(* IEC 61131-3 sources: s7-to-codesys/tests/POUs/Scenarios/FB_Totalizer_ScenarioTest, 7 files *)

(* ---- FB_Totalizer_ScenarioTest.decl.st ---- *)
// AUTO-GENERATED — не редактировать: s7conv gen-tests, сценарии scenarios/FB_Totalizer.csv
// Правка — в CSV (scenarios/README.md), затем python -m s7conv build-corpus.
// Назначение: тесты поведения сконвертированного FB_Totalizer по сценариям CSV (сценариев: 6, строк: 36):
//             один метод-тест на сценарий, строки — по порядку с моделируемым временем GVL_S7Clock.
//             Ожидаемые значения — из CSV (эталонные модели по описанию логики блока), не из
//             результата конвертации.
// Автор:      s7conv 0.1.0 (сгенерировано)
// Версия:     не указана
// Документ:   scenarios/README.md, docs/methodology.md, раздел «Проверка поведения»
FUNCTION_BLOCK FB_Totalizer_ScenarioTest EXTENDS coUnit.FB_TestSuite
VAR
    fbIntegrationAndPulses : FB_Totalizer;  // свой экземпляр на сценарий
    xIntegrationAndPulsesDone : BOOL;  // сценарий выполнен (выполняется один раз)
    fbCutoffAndEnable : FB_Totalizer;  // свой экземпляр на сценарий
    xCutoffAndEnableDone : BOOL;  // сценарий выполнен (выполняется один раз)
    fbResetLevel : FB_Totalizer;  // свой экземпляр на сценарий
    xResetLevelDone : BOOL;  // сценарий выполнен (выполняется один раз)
    fbVariableCycleTime : FB_Totalizer;  // свой экземпляр на сценарий
    xVariableCycleTimeDone : BOOL;  // сценарий выполнен (выполняется один раз)
    fbLargeStepPulsesCatchUp : FB_Totalizer;  // свой экземпляр на сценарий
    xLargeStepPulsesCatchUpDone : BOOL;  // сценарий выполнен (выполняется один раз)
    fbPulseVolumeZero : FB_Totalizer;  // свой экземпляр на сценарий
    xPulseVolumeZeroDone : BOOL;  // сценарий выполнен (выполняется один раз)
END_VAR

(* ---- CutoffAndEnable.method.impl.st ---- *)
// AUTO-GENERATED — не редактировать: scenarios/FB_Totalizer.csv, сценарий CutoffAndEnable
coUnit.TEST('CutoffAndEnable');
IF NOT xCutoffAndEnableDone THEN
    xCutoffAndEnableDone := TRUE;
    GVL_S7Clock.xSimulation := TRUE;

    // #1, t = 0 мс — 0.25 < отсечки 0.5: не считается
    GVL_S7Clock.tSimNow := T#0MS;
    fbCutoffAndEnable.flow := 0.25;
    fbCutoffAndEnable.cycleTime := T#1000MS;
    fbCutoffAndEnable.lowFlowCutoff := 0.5;
    fbCutoffAndEnable.enable := TRUE;
    fbCutoffAndEnable.reset := FALSE;
    fbCutoffAndEnable.pulseVolume := 1.0;
    fbCutoffAndEnable();
    AssertEquals_LREAL(Expected := 0.0,
                       Actual := fbCutoffAndEnable.total,
                       Delta := 0.000001,
                       Message := 'CutoffAndEnable#1 total');
    AssertEquals_LREAL(Expected := 0.0,
                       Actual := fbCutoffAndEnable.lifetimeTotal,
                       Delta := 0.000001,
                       Message := 'CutoffAndEnable#1 lifetimeTotal');
    AssertEquals_DINT(Expected := 0, Actual := fbCutoffAndEnable.pulseCount, Message := 'CutoffAndEnable#1 pulseCount');
    AssertEquals_BOOL(Expected := FALSE, Actual := fbCutoffAndEnable.pulse, Message := 'CutoffAndEnable#1 pulse');
    AssertEquals_BOOL(Expected := TRUE,
                      Actual := fbCutoffAndEnable.cutoffActive,
                      Message := 'CutoffAndEnable#1 cutoffActive');

    // #2, t = 1000 мс — обратный расход ниже отсечки: не считается
    GVL_S7Clock.tSimNow := T#1000MS;
    fbCutoffAndEnable.flow := -10.0;
    fbCutoffAndEnable();
    AssertEquals_LREAL(Expected := 0.0,
                       Actual := fbCutoffAndEnable.total,
                       Delta := 0.000001,
                       Message := 'CutoffAndEnable#2 total');
    AssertEquals_LREAL(Expected := 0.0,
                       Actual := fbCutoffAndEnable.lifetimeTotal,
                       Delta := 0.000001,
                       Message := 'CutoffAndEnable#2 lifetimeTotal');
    AssertEquals_DINT(Expected := 0, Actual := fbCutoffAndEnable.pulseCount, Message := 'CutoffAndEnable#2 pulseCount');
    AssertEquals_BOOL(Expected := FALSE, Actual := fbCutoffAndEnable.pulse, Message := 'CutoffAndEnable#2 pulse');
    AssertEquals_BOOL(Expected := TRUE,
                      Actual := fbCutoffAndEnable.cutoffActive,
                      Message := 'CutoffAndEnable#2 cutoffActive');

    // #3, t = 2000 мс — интегрирование запрещено (отсечка не активна)
    GVL_S7Clock.tSimNow := T#2000MS;
    fbCutoffAndEnable.flow := 450.0;
    fbCutoffAndEnable.enable := FALSE;
    fbCutoffAndEnable();
    AssertEquals_LREAL(Expected := 0.0,
                       Actual := fbCutoffAndEnable.total,
                       Delta := 0.000001,
                       Message := 'CutoffAndEnable#3 total');
    AssertEquals_LREAL(Expected := 0.0,
                       Actual := fbCutoffAndEnable.lifetimeTotal,
                       Delta := 0.000001,
                       Message := 'CutoffAndEnable#3 lifetimeTotal');
    AssertEquals_DINT(Expected := 0, Actual := fbCutoffAndEnable.pulseCount, Message := 'CutoffAndEnable#3 pulseCount');
    AssertEquals_BOOL(Expected := FALSE, Actual := fbCutoffAndEnable.pulse, Message := 'CutoffAndEnable#3 pulse');
    AssertEquals_BOOL(Expected := FALSE,
                      Actual := fbCutoffAndEnable.cutoffActive,
                      Message := 'CutoffAndEnable#3 cutoffActive');

    // #4, t = 3000 мс — разрешено: 0.125 м3
    GVL_S7Clock.tSimNow := T#3000MS;
    fbCutoffAndEnable.enable := TRUE;
    fbCutoffAndEnable();
    AssertEquals_LREAL(Expected := 0.125,
                       Actual := fbCutoffAndEnable.total,
                       Delta := 0.000001,
                       Message := 'CutoffAndEnable#4 total');
    AssertEquals_LREAL(Expected := 0.125,
                       Actual := fbCutoffAndEnable.lifetimeTotal,
                       Delta := 0.000001,
                       Message := 'CutoffAndEnable#4 lifetimeTotal');
    AssertEquals_DINT(Expected := 0, Actual := fbCutoffAndEnable.pulseCount, Message := 'CutoffAndEnable#4 pulseCount');
    AssertEquals_BOOL(Expected := FALSE, Actual := fbCutoffAndEnable.pulse, Message := 'CutoffAndEnable#4 pulse');
    AssertEquals_BOOL(Expected := FALSE,
                      Actual := fbCutoffAndEnable.cutoffActive,
                      Message := 'CutoffAndEnable#4 cutoffActive');

    // #5, t = 4000 мс — 0.5 = отсечке — считается: +0.5/3600 м3
    GVL_S7Clock.tSimNow := T#4000MS;
    fbCutoffAndEnable.flow := 0.5;
    fbCutoffAndEnable();
    AssertEquals_LREAL(Expected := 0.125138889,
                       Actual := fbCutoffAndEnable.total,
                       Delta := 0.000001,
                       Message := 'CutoffAndEnable#5 total');
    AssertEquals_LREAL(Expected := 0.125138889,
                       Actual := fbCutoffAndEnable.lifetimeTotal,
                       Delta := 0.000001,
                       Message := 'CutoffAndEnable#5 lifetimeTotal');
    AssertEquals_DINT(Expected := 0, Actual := fbCutoffAndEnable.pulseCount, Message := 'CutoffAndEnable#5 pulseCount');
    AssertEquals_BOOL(Expected := FALSE, Actual := fbCutoffAndEnable.pulse, Message := 'CutoffAndEnable#5 pulse');
    AssertEquals_BOOL(Expected := FALSE,
                      Actual := fbCutoffAndEnable.cutoffActive,
                      Message := 'CutoffAndEnable#5 cutoffActive');

    // #6, t = 5000 мс — 0.49 < 0.5: не считается
    GVL_S7Clock.tSimNow := T#5000MS;
    fbCutoffAndEnable.flow := 0.49;
    fbCutoffAndEnable();
    AssertEquals_LREAL(Expected := 0.125138889,
                       Actual := fbCutoffAndEnable.total,
                       Delta := 0.000001,
                       Message := 'CutoffAndEnable#6 total');
    AssertEquals_LREAL(Expected := 0.125138889,
                       Actual := fbCutoffAndEnable.lifetimeTotal,
                       Delta := 0.000001,
                       Message := 'CutoffAndEnable#6 lifetimeTotal');
    AssertEquals_DINT(Expected := 0, Actual := fbCutoffAndEnable.pulseCount, Message := 'CutoffAndEnable#6 pulseCount');
    AssertEquals_BOOL(Expected := FALSE, Actual := fbCutoffAndEnable.pulse, Message := 'CutoffAndEnable#6 pulse');
    AssertEquals_BOOL(Expected := TRUE,
                      Actual := fbCutoffAndEnable.cutoffActive,
                      Message := 'CutoffAndEnable#6 cutoffActive');

    GVL_S7Clock.xSimulation := FALSE;
END_IF
coUnit.TEST_FINISHED();

(* ---- IntegrationAndPulses.method.impl.st ---- *)
// AUTO-GENERATED — не редактировать: scenarios/FB_Totalizer.csv, сценарий IntegrationAndPulses
coUnit.TEST('IntegrationAndPulses');
IF NOT xIntegrationAndPulsesDone THEN
    xIntegrationAndPulsesDone := TRUE;
    GVL_S7Clock.xSimulation := TRUE;

    // #1, t = 0 мс — 0.125 м3
    GVL_S7Clock.tSimNow := T#0MS;
    fbIntegrationAndPulses.flow := 450.0;
    fbIntegrationAndPulses.cycleTime := T#1000MS;
    fbIntegrationAndPulses.lowFlowCutoff := 0.5;
    fbIntegrationAndPulses.enable := TRUE;
    fbIntegrationAndPulses.reset := FALSE;
    fbIntegrationAndPulses.pulseVolume := 0.5;
    fbIntegrationAndPulses();
    AssertEquals_LREAL(Expected := 0.125,
                       Actual := fbIntegrationAndPulses.total,
                       Delta := 0.000001,
                       Message := 'IntegrationAndPulses#1 total');
    AssertEquals_LREAL(Expected := 0.125,
                       Actual := fbIntegrationAndPulses.lifetimeTotal,
                       Delta := 0.000001,
                       Message := 'IntegrationAndPulses#1 lifetimeTotal');
    AssertEquals_DINT(Expected := 0,
                      Actual := fbIntegrationAndPulses.pulseCount,
                      Message := 'IntegrationAndPulses#1 pulseCount');
    AssertEquals_BOOL(Expected := FALSE,
                      Actual := fbIntegrationAndPulses.pulse,
                      Message := 'IntegrationAndPulses#1 pulse');
    AssertEquals_BOOL(Expected := FALSE,
                      Actual := fbIntegrationAndPulses.cutoffActive,
                      Message := 'IntegrationAndPulses#1 cutoffActive');

    // #2, t = 1000 мс — 0.25 м3
    GVL_S7Clock.tSimNow := T#1000MS;
    fbIntegrationAndPulses();
    AssertEquals_LREAL(Expected := 0.25,
                       Actual := fbIntegrationAndPulses.total,
                       Delta := 0.000001,
                       Message := 'IntegrationAndPulses#2 total');
    AssertEquals_LREAL(Expected := 0.25,
                       Actual := fbIntegrationAndPulses.lifetimeTotal,
                       Delta := 0.000001,
                       Message := 'IntegrationAndPulses#2 lifetimeTotal');
    AssertEquals_DINT(Expected := 0,
                      Actual := fbIntegrationAndPulses.pulseCount,
                      Message := 'IntegrationAndPulses#2 pulseCount');
    AssertEquals_BOOL(Expected := FALSE,
                      Actual := fbIntegrationAndPulses.pulse,
                      Message := 'IntegrationAndPulses#2 pulse');
    AssertEquals_BOOL(Expected := FALSE,
                      Actual := fbIntegrationAndPulses.cutoffActive,
                      Message := 'IntegrationAndPulses#2 cutoffActive');

    // #3, t = 2000 мс — 0.375 м3
    GVL_S7Clock.tSimNow := T#2000MS;
    fbIntegrationAndPulses();
    AssertEquals_LREAL(Expected := 0.375,
                       Actual := fbIntegrationAndPulses.total,
                       Delta := 0.000001,
                       Message := 'IntegrationAndPulses#3 total');
    AssertEquals_LREAL(Expected := 0.375,
                       Actual := fbIntegrationAndPulses.lifetimeTotal,
                       Delta := 0.000001,
                       Message := 'IntegrationAndPulses#3 lifetimeTotal');
    AssertEquals_DINT(Expected := 0,
                      Actual := fbIntegrationAndPulses.pulseCount,
                      Message := 'IntegrationAndPulses#3 pulseCount');
    AssertEquals_BOOL(Expected := FALSE,
                      Actual := fbIntegrationAndPulses.pulse,
                      Message := 'IntegrationAndPulses#3 pulse');
    AssertEquals_BOOL(Expected := FALSE,
                      Actual := fbIntegrationAndPulses.cutoffActive,
                      Message := 'IntegrationAndPulses#3 cutoffActive');

    // #4, t = 3000 мс — 0.5 м3: импульс №1
    GVL_S7Clock.tSimNow := T#3000MS;
    fbIntegrationAndPulses();
    AssertEquals_LREAL(Expected := 0.5,
                       Actual := fbIntegrationAndPulses.total,
                       Delta := 0.000001,
                       Message := 'IntegrationAndPulses#4 total');
    AssertEquals_LREAL(Expected := 0.5,
                       Actual := fbIntegrationAndPulses.lifetimeTotal,
                       Delta := 0.000001,
                       Message := 'IntegrationAndPulses#4 lifetimeTotal');
    AssertEquals_DINT(Expected := 1,
                      Actual := fbIntegrationAndPulses.pulseCount,
                      Message := 'IntegrationAndPulses#4 pulseCount');
    AssertEquals_BOOL(Expected := TRUE,
                      Actual := fbIntegrationAndPulses.pulse,
                      Message := 'IntegrationAndPulses#4 pulse');
    AssertEquals_BOOL(Expected := FALSE,
                      Actual := fbIntegrationAndPulses.cutoffActive,
                      Message := 'IntegrationAndPulses#4 cutoffActive');

    // #5, t = 4000 мс — 0.625 м3, импульса нет
    GVL_S7Clock.tSimNow := T#4000MS;
    fbIntegrationAndPulses();
    AssertEquals_LREAL(Expected := 0.625,
                       Actual := fbIntegrationAndPulses.total,
                       Delta := 0.000001,
                       Message := 'IntegrationAndPulses#5 total');
    AssertEquals_LREAL(Expected := 0.625,
                       Actual := fbIntegrationAndPulses.lifetimeTotal,
                       Delta := 0.000001,
                       Message := 'IntegrationAndPulses#5 lifetimeTotal');
    AssertEquals_DINT(Expected := 1,
                      Actual := fbIntegrationAndPulses.pulseCount,
                      Message := 'IntegrationAndPulses#5 pulseCount');
    AssertEquals_BOOL(Expected := FALSE,
                      Actual := fbIntegrationAndPulses.pulse,
                      Message := 'IntegrationAndPulses#5 pulse');
    AssertEquals_BOOL(Expected := FALSE,
                      Actual := fbIntegrationAndPulses.cutoffActive,
                      Message := 'IntegrationAndPulses#5 cutoffActive');

    // #6, t = 5000 мс — 0.75 м3
    GVL_S7Clock.tSimNow := T#5000MS;
    fbIntegrationAndPulses();
    AssertEquals_LREAL(Expected := 0.75,
                       Actual := fbIntegrationAndPulses.total,
                       Delta := 0.000001,
                       Message := 'IntegrationAndPulses#6 total');
    AssertEquals_LREAL(Expected := 0.75,
                       Actual := fbIntegrationAndPulses.lifetimeTotal,
                       Delta := 0.000001,
                       Message := 'IntegrationAndPulses#6 lifetimeTotal');
    AssertEquals_DINT(Expected := 1,
                      Actual := fbIntegrationAndPulses.pulseCount,
                      Message := 'IntegrationAndPulses#6 pulseCount');
    AssertEquals_BOOL(Expected := FALSE,
                      Actual := fbIntegrationAndPulses.pulse,
                      Message := 'IntegrationAndPulses#6 pulse');
    AssertEquals_BOOL(Expected := FALSE,
                      Actual := fbIntegrationAndPulses.cutoffActive,
                      Message := 'IntegrationAndPulses#6 cutoffActive');

    // #7, t = 6000 мс — 0.875 м3
    GVL_S7Clock.tSimNow := T#6000MS;
    fbIntegrationAndPulses();
    AssertEquals_LREAL(Expected := 0.875,
                       Actual := fbIntegrationAndPulses.total,
                       Delta := 0.000001,
                       Message := 'IntegrationAndPulses#7 total');
    AssertEquals_LREAL(Expected := 0.875,
                       Actual := fbIntegrationAndPulses.lifetimeTotal,
                       Delta := 0.000001,
                       Message := 'IntegrationAndPulses#7 lifetimeTotal');
    AssertEquals_DINT(Expected := 1,
                      Actual := fbIntegrationAndPulses.pulseCount,
                      Message := 'IntegrationAndPulses#7 pulseCount');
    AssertEquals_BOOL(Expected := FALSE,
                      Actual := fbIntegrationAndPulses.pulse,
                      Message := 'IntegrationAndPulses#7 pulse');
    AssertEquals_BOOL(Expected := FALSE,
                      Actual := fbIntegrationAndPulses.cutoffActive,
                      Message := 'IntegrationAndPulses#7 cutoffActive');

    // #8, t = 7000 мс — 1.0 м3: импульс №2
    GVL_S7Clock.tSimNow := T#7000MS;
    fbIntegrationAndPulses();
    AssertEquals_LREAL(Expected := 1.0,
                       Actual := fbIntegrationAndPulses.total,
                       Delta := 0.000001,
                       Message := 'IntegrationAndPulses#8 total');
    AssertEquals_LREAL(Expected := 1.0,
                       Actual := fbIntegrationAndPulses.lifetimeTotal,
                       Delta := 0.000001,
                       Message := 'IntegrationAndPulses#8 lifetimeTotal');
    AssertEquals_DINT(Expected := 2,
                      Actual := fbIntegrationAndPulses.pulseCount,
                      Message := 'IntegrationAndPulses#8 pulseCount');
    AssertEquals_BOOL(Expected := TRUE,
                      Actual := fbIntegrationAndPulses.pulse,
                      Message := 'IntegrationAndPulses#8 pulse');
    AssertEquals_BOOL(Expected := FALSE,
                      Actual := fbIntegrationAndPulses.cutoffActive,
                      Message := 'IntegrationAndPulses#8 cutoffActive');

    // #9, t = 8000 мс — 900 м3/ч: +0.25 м3 = 1.25
    GVL_S7Clock.tSimNow := T#8000MS;
    fbIntegrationAndPulses.flow := 900.0;
    fbIntegrationAndPulses();
    AssertEquals_LREAL(Expected := 1.25,
                       Actual := fbIntegrationAndPulses.total,
                       Delta := 0.000001,
                       Message := 'IntegrationAndPulses#9 total');
    AssertEquals_LREAL(Expected := 1.25,
                       Actual := fbIntegrationAndPulses.lifetimeTotal,
                       Delta := 0.000001,
                       Message := 'IntegrationAndPulses#9 lifetimeTotal');
    AssertEquals_DINT(Expected := 2,
                      Actual := fbIntegrationAndPulses.pulseCount,
                      Message := 'IntegrationAndPulses#9 pulseCount');
    AssertEquals_BOOL(Expected := FALSE,
                      Actual := fbIntegrationAndPulses.pulse,
                      Message := 'IntegrationAndPulses#9 pulse');
    AssertEquals_BOOL(Expected := FALSE,
                      Actual := fbIntegrationAndPulses.cutoffActive,
                      Message := 'IntegrationAndPulses#9 cutoffActive');

    // #10, t = 9000 мс — 1.5 м3: импульс №3
    GVL_S7Clock.tSimNow := T#9000MS;
    fbIntegrationAndPulses();
    AssertEquals_LREAL(Expected := 1.5,
                       Actual := fbIntegrationAndPulses.total,
                       Delta := 0.000001,
                       Message := 'IntegrationAndPulses#10 total');
    AssertEquals_LREAL(Expected := 1.5,
                       Actual := fbIntegrationAndPulses.lifetimeTotal,
                       Delta := 0.000001,
                       Message := 'IntegrationAndPulses#10 lifetimeTotal');
    AssertEquals_DINT(Expected := 3,
                      Actual := fbIntegrationAndPulses.pulseCount,
                      Message := 'IntegrationAndPulses#10 pulseCount');
    AssertEquals_BOOL(Expected := TRUE,
                      Actual := fbIntegrationAndPulses.pulse,
                      Message := 'IntegrationAndPulses#10 pulse');
    AssertEquals_BOOL(Expected := FALSE,
                      Actual := fbIntegrationAndPulses.cutoffActive,
                      Message := 'IntegrationAndPulses#10 cutoffActive');

    GVL_S7Clock.xSimulation := FALSE;
END_IF
coUnit.TEST_FINISHED();

(* ---- LargeStepPulsesCatchUp.method.impl.st ---- *)
// AUTO-GENERATED — не редактировать: scenarios/FB_Totalizer.csv, сценарий LargeStepPulsesCatchUp
coUnit.TEST('LargeStepPulsesCatchUp');
IF NOT xLargeStepPulsesCatchUpDone THEN
    xLargeStepPulsesCatchUpDone := TRUE;
    GVL_S7Clock.xSimulation := TRUE;

    // #1, t = 0 мс — +1.0 м3 за вызов: импульс №1, остаток 0.5
    GVL_S7Clock.tSimNow := T#0MS;
    fbLargeStepPulsesCatchUp.flow := 3600.0;
    fbLargeStepPulsesCatchUp.cycleTime := T#1000MS;
    fbLargeStepPulsesCatchUp.lowFlowCutoff := 0.5;
    fbLargeStepPulsesCatchUp.enable := TRUE;
    fbLargeStepPulsesCatchUp.reset := FALSE;
    fbLargeStepPulsesCatchUp.pulseVolume := 0.5;
    fbLargeStepPulsesCatchUp();
    AssertEquals_LREAL(Expected := 1.0,
                       Actual := fbLargeStepPulsesCatchUp.total,
                       Delta := 0.000001,
                       Message := 'LargeStepPulsesCatchUp#1 total');
    AssertEquals_LREAL(Expected := 1.0,
                       Actual := fbLargeStepPulsesCatchUp.lifetimeTotal,
                       Delta := 0.000001,
                       Message := 'LargeStepPulsesCatchUp#1 lifetimeTotal');
    AssertEquals_DINT(Expected := 1,
                      Actual := fbLargeStepPulsesCatchUp.pulseCount,
                      Message := 'LargeStepPulsesCatchUp#1 pulseCount');
    AssertEquals_BOOL(Expected := TRUE,
                      Actual := fbLargeStepPulsesCatchUp.pulse,
                      Message := 'LargeStepPulsesCatchUp#1 pulse');
    AssertEquals_BOOL(Expected := FALSE,
                      Actual := fbLargeStepPulsesCatchUp.cutoffActive,
                      Message := 'LargeStepPulsesCatchUp#1 cutoffActive');

    // #2, t = 1000 мс — 2.0 м3: импульс №2, остаток 1.0
    GVL_S7Clock.tSimNow := T#1000MS;
    fbLargeStepPulsesCatchUp();
    AssertEquals_LREAL(Expected := 2.0,
                       Actual := fbLargeStepPulsesCatchUp.total,
                       Delta := 0.000001,
                       Message := 'LargeStepPulsesCatchUp#2 total');
    AssertEquals_LREAL(Expected := 2.0,
                       Actual := fbLargeStepPulsesCatchUp.lifetimeTotal,
                       Delta := 0.000001,
                       Message := 'LargeStepPulsesCatchUp#2 lifetimeTotal');
    AssertEquals_DINT(Expected := 2,
                      Actual := fbLargeStepPulsesCatchUp.pulseCount,
                      Message := 'LargeStepPulsesCatchUp#2 pulseCount');
    AssertEquals_BOOL(Expected := TRUE,
                      Actual := fbLargeStepPulsesCatchUp.pulse,
                      Message := 'LargeStepPulsesCatchUp#2 pulse');
    AssertEquals_BOOL(Expected := FALSE,
                      Actual := fbLargeStepPulsesCatchUp.cutoffActive,
                      Message := 'LargeStepPulsesCatchUp#2 cutoffActive');

    // #3, t = 2000 мс — расход 0: импульс №3 из остатка, остаток 0.5
    GVL_S7Clock.tSimNow := T#2000MS;
    fbLargeStepPulsesCatchUp.flow := 0.0;
    fbLargeStepPulsesCatchUp();
    AssertEquals_LREAL(Expected := 2.0,
                       Actual := fbLargeStepPulsesCatchUp.total,
                       Delta := 0.000001,
                       Message := 'LargeStepPulsesCatchUp#3 total');
    AssertEquals_LREAL(Expected := 2.0,
                       Actual := fbLargeStepPulsesCatchUp.lifetimeTotal,
                       Delta := 0.000001,
                       Message := 'LargeStepPulsesCatchUp#3 lifetimeTotal');
    AssertEquals_DINT(Expected := 3,
                      Actual := fbLargeStepPulsesCatchUp.pulseCount,
                      Message := 'LargeStepPulsesCatchUp#3 pulseCount');
    AssertEquals_BOOL(Expected := TRUE,
                      Actual := fbLargeStepPulsesCatchUp.pulse,
                      Message := 'LargeStepPulsesCatchUp#3 pulse');
    AssertEquals_BOOL(Expected := TRUE,
                      Actual := fbLargeStepPulsesCatchUp.cutoffActive,
                      Message := 'LargeStepPulsesCatchUp#3 cutoffActive');

    // #4, t = 3000 мс — импульс №4, остаток 0
    GVL_S7Clock.tSimNow := T#3000MS;
    fbLargeStepPulsesCatchUp();
    AssertEquals_LREAL(Expected := 2.0,
                       Actual := fbLargeStepPulsesCatchUp.total,
                       Delta := 0.000001,
                       Message := 'LargeStepPulsesCatchUp#4 total');
    AssertEquals_LREAL(Expected := 2.0,
                       Actual := fbLargeStepPulsesCatchUp.lifetimeTotal,
                       Delta := 0.000001,
                       Message := 'LargeStepPulsesCatchUp#4 lifetimeTotal');
    AssertEquals_DINT(Expected := 4,
                      Actual := fbLargeStepPulsesCatchUp.pulseCount,
                      Message := 'LargeStepPulsesCatchUp#4 pulseCount');
    AssertEquals_BOOL(Expected := TRUE,
                      Actual := fbLargeStepPulsesCatchUp.pulse,
                      Message := 'LargeStepPulsesCatchUp#4 pulse');
    AssertEquals_BOOL(Expected := TRUE,
                      Actual := fbLargeStepPulsesCatchUp.cutoffActive,
                      Message := 'LargeStepPulsesCatchUp#4 cutoffActive');

    // #5, t = 4000 мс — импульсов нет: 4 x 0.5 = 2.0 м3
    GVL_S7Clock.tSimNow := T#4000MS;
    fbLargeStepPulsesCatchUp();
    AssertEquals_LREAL(Expected := 2.0,
                       Actual := fbLargeStepPulsesCatchUp.total,
                       Delta := 0.000001,
                       Message := 'LargeStepPulsesCatchUp#5 total');
    AssertEquals_LREAL(Expected := 2.0,
                       Actual := fbLargeStepPulsesCatchUp.lifetimeTotal,
                       Delta := 0.000001,
                       Message := 'LargeStepPulsesCatchUp#5 lifetimeTotal');
    AssertEquals_DINT(Expected := 4,
                      Actual := fbLargeStepPulsesCatchUp.pulseCount,
                      Message := 'LargeStepPulsesCatchUp#5 pulseCount');
    AssertEquals_BOOL(Expected := FALSE,
                      Actual := fbLargeStepPulsesCatchUp.pulse,
                      Message := 'LargeStepPulsesCatchUp#5 pulse');
    AssertEquals_BOOL(Expected := TRUE,
                      Actual := fbLargeStepPulsesCatchUp.cutoffActive,
                      Message := 'LargeStepPulsesCatchUp#5 cutoffActive');

    GVL_S7Clock.xSimulation := FALSE;
END_IF
coUnit.TEST_FINISHED();

(* ---- PulseVolumeZero.method.impl.st ---- *)
// AUTO-GENERATED — не редактировать: scenarios/FB_Totalizer.csv, сценарий PulseVolumeZero
coUnit.TEST('PulseVolumeZero');
IF NOT xPulseVolumeZeroDone THEN
    xPulseVolumeZeroDone := TRUE;
    GVL_S7Clock.xSimulation := TRUE;

    // #1, t = 0 мс — 1.0 м3, импульсов нет
    GVL_S7Clock.tSimNow := T#0MS;
    fbPulseVolumeZero.flow := 3600.0;
    fbPulseVolumeZero.cycleTime := T#1000MS;
    fbPulseVolumeZero.lowFlowCutoff := 0.5;
    fbPulseVolumeZero.enable := TRUE;
    fbPulseVolumeZero.reset := FALSE;
    fbPulseVolumeZero.pulseVolume := 0.0;
    fbPulseVolumeZero();
    AssertEquals_LREAL(Expected := 1.0,
                       Actual := fbPulseVolumeZero.total,
                       Delta := 0.000001,
                       Message := 'PulseVolumeZero#1 total');
    AssertEquals_LREAL(Expected := 1.0,
                       Actual := fbPulseVolumeZero.lifetimeTotal,
                       Delta := 0.000001,
                       Message := 'PulseVolumeZero#1 lifetimeTotal');
    AssertEquals_DINT(Expected := 0, Actual := fbPulseVolumeZero.pulseCount, Message := 'PulseVolumeZero#1 pulseCount');
    AssertEquals_BOOL(Expected := FALSE, Actual := fbPulseVolumeZero.pulse, Message := 'PulseVolumeZero#1 pulse');
    AssertEquals_BOOL(Expected := FALSE,
                      Actual := fbPulseVolumeZero.cutoffActive,
                      Message := 'PulseVolumeZero#1 cutoffActive');

    // #2, t = 1000 мс — 2.0 м3, импульсов нет
    GVL_S7Clock.tSimNow := T#1000MS;
    fbPulseVolumeZero();
    AssertEquals_LREAL(Expected := 2.0,
                       Actual := fbPulseVolumeZero.total,
                       Delta := 0.000001,
                       Message := 'PulseVolumeZero#2 total');
    AssertEquals_LREAL(Expected := 2.0,
                       Actual := fbPulseVolumeZero.lifetimeTotal,
                       Delta := 0.000001,
                       Message := 'PulseVolumeZero#2 lifetimeTotal');
    AssertEquals_DINT(Expected := 0, Actual := fbPulseVolumeZero.pulseCount, Message := 'PulseVolumeZero#2 pulseCount');
    AssertEquals_BOOL(Expected := FALSE, Actual := fbPulseVolumeZero.pulse, Message := 'PulseVolumeZero#2 pulse');
    AssertEquals_BOOL(Expected := FALSE,
                      Actual := fbPulseVolumeZero.cutoffActive,
                      Message := 'PulseVolumeZero#2 cutoffActive');

    GVL_S7Clock.xSimulation := FALSE;
END_IF
coUnit.TEST_FINISHED();

(* ---- ResetLevel.method.impl.st ---- *)
// AUTO-GENERATED — не редактировать: scenarios/FB_Totalizer.csv, сценарий ResetLevel
coUnit.TEST('ResetLevel');
IF NOT xResetLevelDone THEN
    xResetLevelDone := TRUE;
    GVL_S7Clock.xSimulation := TRUE;

    // #1, t = 0 мс — 0.25 м3
    GVL_S7Clock.tSimNow := T#0MS;
    fbResetLevel.flow := 900.0;
    fbResetLevel.cycleTime := T#1000MS;
    fbResetLevel.lowFlowCutoff := 0.5;
    fbResetLevel.enable := TRUE;
    fbResetLevel.reset := FALSE;
    fbResetLevel.pulseVolume := 1.0;
    fbResetLevel();
    AssertEquals_LREAL(Expected := 0.25,
                       Actual := fbResetLevel.total,
                       Delta := 0.000001,
                       Message := 'ResetLevel#1 total');
    AssertEquals_LREAL(Expected := 0.25,
                       Actual := fbResetLevel.lifetimeTotal,
                       Delta := 0.000001,
                       Message := 'ResetLevel#1 lifetimeTotal');
    AssertEquals_DINT(Expected := 0, Actual := fbResetLevel.pulseCount, Message := 'ResetLevel#1 pulseCount');
    AssertEquals_BOOL(Expected := FALSE, Actual := fbResetLevel.pulse, Message := 'ResetLevel#1 pulse');
    AssertEquals_BOOL(Expected := FALSE, Actual := fbResetLevel.cutoffActive, Message := 'ResetLevel#1 cutoffActive');

    // #2, t = 1000 мс — 0.5 м3
    GVL_S7Clock.tSimNow := T#1000MS;
    fbResetLevel();
    AssertEquals_LREAL(Expected := 0.5,
                       Actual := fbResetLevel.total,
                       Delta := 0.000001,
                       Message := 'ResetLevel#2 total');
    AssertEquals_LREAL(Expected := 0.5,
                       Actual := fbResetLevel.lifetimeTotal,
                       Delta := 0.000001,
                       Message := 'ResetLevel#2 lifetimeTotal');
    AssertEquals_DINT(Expected := 0, Actual := fbResetLevel.pulseCount, Message := 'ResetLevel#2 pulseCount');
    AssertEquals_BOOL(Expected := FALSE, Actual := fbResetLevel.pulse, Message := 'ResetLevel#2 pulse');
    AssertEquals_BOOL(Expected := FALSE, Actual := fbResetLevel.cutoffActive, Message := 'ResetLevel#2 cutoffActive');

    // #3, t = 2000 мс — сброс: total 0, общий 0.75
    GVL_S7Clock.tSimNow := T#2000MS;
    fbResetLevel.reset := TRUE;
    fbResetLevel();
    AssertEquals_LREAL(Expected := 0.0,
                       Actual := fbResetLevel.total,
                       Delta := 0.000001,
                       Message := 'ResetLevel#3 total');
    AssertEquals_LREAL(Expected := 0.75,
                       Actual := fbResetLevel.lifetimeTotal,
                       Delta := 0.000001,
                       Message := 'ResetLevel#3 lifetimeTotal');
    AssertEquals_DINT(Expected := 0, Actual := fbResetLevel.pulseCount, Message := 'ResetLevel#3 pulseCount');
    AssertEquals_BOOL(Expected := FALSE, Actual := fbResetLevel.pulse, Message := 'ResetLevel#3 pulse');
    AssertEquals_BOOL(Expected := FALSE, Actual := fbResetLevel.cutoffActive, Message := 'ResetLevel#3 cutoffActive');

    // #4, t = 3000 мс — сброс держится: total 0, общий 1.0
    GVL_S7Clock.tSimNow := T#3000MS;
    fbResetLevel();
    AssertEquals_LREAL(Expected := 0.0,
                       Actual := fbResetLevel.total,
                       Delta := 0.000001,
                       Message := 'ResetLevel#4 total');
    AssertEquals_LREAL(Expected := 1.0,
                       Actual := fbResetLevel.lifetimeTotal,
                       Delta := 0.000001,
                       Message := 'ResetLevel#4 lifetimeTotal');
    AssertEquals_DINT(Expected := 0, Actual := fbResetLevel.pulseCount, Message := 'ResetLevel#4 pulseCount');
    AssertEquals_BOOL(Expected := FALSE, Actual := fbResetLevel.pulse, Message := 'ResetLevel#4 pulse');
    AssertEquals_BOOL(Expected := FALSE, Actual := fbResetLevel.cutoffActive, Message := 'ResetLevel#4 cutoffActive');

    // #5, t = 4000 мс — сброс снят: total 0.25, общий 1.25
    GVL_S7Clock.tSimNow := T#4000MS;
    fbResetLevel.reset := FALSE;
    fbResetLevel();
    AssertEquals_LREAL(Expected := 0.25,
                       Actual := fbResetLevel.total,
                       Delta := 0.000001,
                       Message := 'ResetLevel#5 total');
    AssertEquals_LREAL(Expected := 1.25,
                       Actual := fbResetLevel.lifetimeTotal,
                       Delta := 0.000001,
                       Message := 'ResetLevel#5 lifetimeTotal');
    AssertEquals_DINT(Expected := 0, Actual := fbResetLevel.pulseCount, Message := 'ResetLevel#5 pulseCount');
    AssertEquals_BOOL(Expected := FALSE, Actual := fbResetLevel.pulse, Message := 'ResetLevel#5 pulse');
    AssertEquals_BOOL(Expected := FALSE, Actual := fbResetLevel.cutoffActive, Message := 'ResetLevel#5 cutoffActive');

    // #6, t = 5000 мс — 0.5
    GVL_S7Clock.tSimNow := T#5000MS;
    fbResetLevel();
    AssertEquals_LREAL(Expected := 0.5,
                       Actual := fbResetLevel.total,
                       Delta := 0.000001,
                       Message := 'ResetLevel#6 total');
    AssertEquals_LREAL(Expected := 1.5,
                       Actual := fbResetLevel.lifetimeTotal,
                       Delta := 0.000001,
                       Message := 'ResetLevel#6 lifetimeTotal');
    AssertEquals_DINT(Expected := 0, Actual := fbResetLevel.pulseCount, Message := 'ResetLevel#6 pulseCount');
    AssertEquals_BOOL(Expected := FALSE, Actual := fbResetLevel.pulse, Message := 'ResetLevel#6 pulse');
    AssertEquals_BOOL(Expected := FALSE, Actual := fbResetLevel.cutoffActive, Message := 'ResetLevel#6 cutoffActive');

    // #7, t = 6000 мс — 0.75
    GVL_S7Clock.tSimNow := T#6000MS;
    fbResetLevel();
    AssertEquals_LREAL(Expected := 0.75,
                       Actual := fbResetLevel.total,
                       Delta := 0.000001,
                       Message := 'ResetLevel#7 total');
    AssertEquals_LREAL(Expected := 1.75,
                       Actual := fbResetLevel.lifetimeTotal,
                       Delta := 0.000001,
                       Message := 'ResetLevel#7 lifetimeTotal');
    AssertEquals_DINT(Expected := 0, Actual := fbResetLevel.pulseCount, Message := 'ResetLevel#7 pulseCount');
    AssertEquals_BOOL(Expected := FALSE, Actual := fbResetLevel.pulse, Message := 'ResetLevel#7 pulse');
    AssertEquals_BOOL(Expected := FALSE, Actual := fbResetLevel.cutoffActive, Message := 'ResetLevel#7 cutoffActive');

    // #8, t = 7000 мс — 1.0 м3 после сброса: импульс №1
    GVL_S7Clock.tSimNow := T#7000MS;
    fbResetLevel();
    AssertEquals_LREAL(Expected := 1.0,
                       Actual := fbResetLevel.total,
                       Delta := 0.000001,
                       Message := 'ResetLevel#8 total');
    AssertEquals_LREAL(Expected := 2.0,
                       Actual := fbResetLevel.lifetimeTotal,
                       Delta := 0.000001,
                       Message := 'ResetLevel#8 lifetimeTotal');
    AssertEquals_DINT(Expected := 1, Actual := fbResetLevel.pulseCount, Message := 'ResetLevel#8 pulseCount');
    AssertEquals_BOOL(Expected := TRUE, Actual := fbResetLevel.pulse, Message := 'ResetLevel#8 pulse');
    AssertEquals_BOOL(Expected := FALSE, Actual := fbResetLevel.cutoffActive, Message := 'ResetLevel#8 cutoffActive');

    GVL_S7Clock.xSimulation := FALSE;
END_IF
coUnit.TEST_FINISHED();

(* ---- VariableCycleTime.method.impl.st ---- *)
// AUTO-GENERATED — не редактировать: scenarios/FB_Totalizer.csv, сценарий VariableCycleTime
coUnit.TEST('VariableCycleTime');
IF NOT xVariableCycleTimeDone THEN
    xVariableCycleTimeDone := TRUE;
    GVL_S7Clock.xSimulation := TRUE;

    // #1, t = 0 мс — 0.5 с: 0.0625 м3
    GVL_S7Clock.tSimNow := T#0MS;
    fbVariableCycleTime.flow := 450.0;
    fbVariableCycleTime.cycleTime := T#500MS;
    fbVariableCycleTime.lowFlowCutoff := 0.5;
    fbVariableCycleTime.enable := TRUE;
    fbVariableCycleTime.reset := FALSE;
    fbVariableCycleTime.pulseVolume := 0.5;
    fbVariableCycleTime();
    AssertEquals_LREAL(Expected := 0.0625,
                       Actual := fbVariableCycleTime.total,
                       Delta := 0.000001,
                       Message := 'VariableCycleTime#1 total');
    AssertEquals_LREAL(Expected := 0.0625,
                       Actual := fbVariableCycleTime.lifetimeTotal,
                       Delta := 0.000001,
                       Message := 'VariableCycleTime#1 lifetimeTotal');
    AssertEquals_DINT(Expected := 0,
                      Actual := fbVariableCycleTime.pulseCount,
                      Message := 'VariableCycleTime#1 pulseCount');
    AssertEquals_BOOL(Expected := FALSE, Actual := fbVariableCycleTime.pulse, Message := 'VariableCycleTime#1 pulse');
    AssertEquals_BOOL(Expected := FALSE,
                      Actual := fbVariableCycleTime.cutoffActive,
                      Message := 'VariableCycleTime#1 cutoffActive');

    // #2, t = 500 мс — 0.125 м3
    GVL_S7Clock.tSimNow := T#500MS;
    fbVariableCycleTime();
    AssertEquals_LREAL(Expected := 0.125,
                       Actual := fbVariableCycleTime.total,
                       Delta := 0.000001,
                       Message := 'VariableCycleTime#2 total');
    AssertEquals_LREAL(Expected := 0.125,
                       Actual := fbVariableCycleTime.lifetimeTotal,
                       Delta := 0.000001,
                       Message := 'VariableCycleTime#2 lifetimeTotal');
    AssertEquals_DINT(Expected := 0,
                      Actual := fbVariableCycleTime.pulseCount,
                      Message := 'VariableCycleTime#2 pulseCount');
    AssertEquals_BOOL(Expected := FALSE, Actual := fbVariableCycleTime.pulse, Message := 'VariableCycleTime#2 pulse');
    AssertEquals_BOOL(Expected := FALSE,
                      Actual := fbVariableCycleTime.cutoffActive,
                      Message := 'VariableCycleTime#2 cutoffActive');

    // #3, t = 2500 мс — 2 с: +0.25 = 0.375 м3
    GVL_S7Clock.tSimNow := T#2500MS;
    fbVariableCycleTime.cycleTime := T#2000MS;
    fbVariableCycleTime();
    AssertEquals_LREAL(Expected := 0.375,
                       Actual := fbVariableCycleTime.total,
                       Delta := 0.000001,
                       Message := 'VariableCycleTime#3 total');
    AssertEquals_LREAL(Expected := 0.375,
                       Actual := fbVariableCycleTime.lifetimeTotal,
                       Delta := 0.000001,
                       Message := 'VariableCycleTime#3 lifetimeTotal');
    AssertEquals_DINT(Expected := 0,
                      Actual := fbVariableCycleTime.pulseCount,
                      Message := 'VariableCycleTime#3 pulseCount');
    AssertEquals_BOOL(Expected := FALSE, Actual := fbVariableCycleTime.pulse, Message := 'VariableCycleTime#3 pulse');
    AssertEquals_BOOL(Expected := FALSE,
                      Actual := fbVariableCycleTime.cutoffActive,
                      Message := 'VariableCycleTime#3 cutoffActive');

    // #4, t = 2600 мс — 0.1 с: +0.0125 = 0.3875 м3
    GVL_S7Clock.tSimNow := T#2600MS;
    fbVariableCycleTime.cycleTime := T#100MS;
    fbVariableCycleTime();
    AssertEquals_LREAL(Expected := 0.3875,
                       Actual := fbVariableCycleTime.total,
                       Delta := 0.000001,
                       Message := 'VariableCycleTime#4 total');
    AssertEquals_LREAL(Expected := 0.3875,
                       Actual := fbVariableCycleTime.lifetimeTotal,
                       Delta := 0.000001,
                       Message := 'VariableCycleTime#4 lifetimeTotal');
    AssertEquals_DINT(Expected := 0,
                      Actual := fbVariableCycleTime.pulseCount,
                      Message := 'VariableCycleTime#4 pulseCount');
    AssertEquals_BOOL(Expected := FALSE, Actual := fbVariableCycleTime.pulse, Message := 'VariableCycleTime#4 pulse');
    AssertEquals_BOOL(Expected := FALSE,
                      Actual := fbVariableCycleTime.cutoffActive,
                      Message := 'VariableCycleTime#4 cutoffActive');

    // #5, t = 2700 мс — 0.4 м3, до импульса 0.1 м3
    GVL_S7Clock.tSimNow := T#2700MS;
    fbVariableCycleTime();
    AssertEquals_LREAL(Expected := 0.4,
                       Actual := fbVariableCycleTime.total,
                       Delta := 0.000001,
                       Message := 'VariableCycleTime#5 total');
    AssertEquals_LREAL(Expected := 0.4,
                       Actual := fbVariableCycleTime.lifetimeTotal,
                       Delta := 0.000001,
                       Message := 'VariableCycleTime#5 lifetimeTotal');
    AssertEquals_DINT(Expected := 0,
                      Actual := fbVariableCycleTime.pulseCount,
                      Message := 'VariableCycleTime#5 pulseCount');
    AssertEquals_BOOL(Expected := FALSE, Actual := fbVariableCycleTime.pulse, Message := 'VariableCycleTime#5 pulse');
    AssertEquals_BOOL(Expected := FALSE,
                      Actual := fbVariableCycleTime.cutoffActive,
                      Message := 'VariableCycleTime#5 cutoffActive');

    GVL_S7Clock.xSimulation := FALSE;
END_IF
coUnit.TEST_FINISHED();
